(* IEC 61131-3 sources: avi-aoi-management/scripts/ai-eval/ngau-nhien/lib/st-scl/mau-scl/st-ud7-van-hai-cuon/src, 2 files *)

(* ---- ViTriVan.st ---- *)
FUNCTION "ViTriVan" : Int
{ S7_Optimized_Access := 'TRUE' }
VERSION : 0.1
   VAR_INPUT
      CT_MO : Bool;
      CT_DONG : Bool;
   END_VAR

   REGION Giai ma vi tri van
      IF #CT_MO AND #CT_DONG THEN
         #ViTriVan := 3;
      ELSIF #CT_MO THEN
         #ViTriVan := 1;
      ELSIF #CT_DONG THEN
         #ViTriVan := 2;
      ELSE
         #ViTriVan := 0;
      END_IF;
   END_REGION
END_FUNCTION

(* ---- VanHaiCuon.st ---- *)
FUNCTION_BLOCK "VanHaiCuon"
{ S7_Optimized_Access := 'TRUE' }
VERSION : 0.1
   VAR_INPUT
      MO : Bool;
      DONG : Bool;
      CT_MO : Bool;
      CT_DONG : Bool;
      RESET : Bool;
      T_HANH_TRINH : Time;
   END_VAR

   VAR_OUTPUT
      CUON_MO : Bool;
      CUON_DONG : Bool;
      TRANG_THAI : Int;  // 1 DANG_MO, 2 DANG_DONG, 3 DA_MO, 4 DA_DONG, 5 GIUA_CHUNG, 9 LOI
      MA_LOI : Int;      // 0, 1 hành trình, 2 công tắc
   END_VAR

   VAR
      rtMo : R_TRIG;
      rtDong : R_TRIG;
      tBuoc : TON_TIME;       // ET = thời gian đã ở bước hiện tại
      tt : Int;          // 0 NGHI, 1 CHAY_MO, 2 CHAY_DONG, 3 DAO_MO, 4 DAO_DONG, 9 LOI
      ttTruoc : Int;
   END_VAR

   VAR_TEMP
      vt : Int;
      eMo : Bool;
      eDong : Bool;
   END_VAR

   REGION Cam bien va suon lenh
      #vt := "ViTriVan"(CT_MO := #CT_MO, CT_DONG := #CT_DONG);
      #rtMo(CLK := #MO);
      #rtDong(CLK := #DONG);
      #eMo := #rtMo.Q AND NOT #rtDong.Q;
      #eDong := #rtDong.Q AND NOT #rtMo.Q;
      #tBuoc(IN := TRUE, PT := T#24h);
   END_REGION

   REGION May trang thai
      IF #vt = 3 THEN
         IF #tt <> 9 THEN #MA_LOI := 2; END_IF;
         #tt := 9;
      ELSE
         CASE #tt OF
            0:
               IF #eMo AND #vt <> 1 THEN #tt := 1;
               ELSIF #eDong AND #vt <> 2 THEN #tt := 2;
               END_IF;
            1:
               IF #vt = 1 THEN #tt := 0;
               ELSIF #eDong THEN #tt := 4;
               ELSIF #tBuoc.ET >= #T_HANH_TRINH THEN #tt := 9; #MA_LOI := 1;
               END_IF;
            2:
               IF #vt = 2 THEN #tt := 0;
               ELSIF #eMo THEN #tt := 3;
               ELSIF #tBuoc.ET >= #T_HANH_TRINH THEN #tt := 9; #MA_LOI := 1;
               END_IF;
            3: #tt := 1;
            4: #tt := 2;
            9:
               IF #RESET THEN #tt := 0; #MA_LOI := 0; END_IF;
         END_CASE;
      END_IF;
      IF #tt <> #ttTruoc THEN
         #tBuoc(IN := FALSE);
         #tBuoc(IN := TRUE, PT := T#24h);
      END_IF;
      #ttTruoc := #tt;
   END_REGION

   REGION Dau ra
      #CUON_MO := #tt = 1;
      #CUON_DONG := #tt = 2;
      CASE #tt OF
         1, 3: #TRANG_THAI := 1;
         2, 4: #TRANG_THAI := 2;
         9: #TRANG_THAI := 9;
         ELSE
            IF #vt = 1 THEN #TRANG_THAI := 3;
            ELSIF #vt = 2 THEN #TRANG_THAI := 4;
            ELSE #TRANG_THAI := 5;
            END_IF;
      END_CASE;
   END_REGION
END_FUNCTION_BLOCK
